(* IEC 61131-3 sources: nautilus/tools/blackbox/projects/2026-10-24-001d/typed, 2 files *)

(* ---- types.st ---- *)
(* library file: types used by the typed project *)
TYPE Mode : (Idle, Run := 10, Fault) := Idle; END_TYPE
TYPE Drive : STRUCT
    Speed : REAL;
    Amps  : REAL;
  END_STRUCT;
END_TYPE
TYPE Motor : STRUCT
    Running : BOOL;
    Fault   : BOOL;
    Starts  : DINT;
    Drive   : Drive;
    State   : Mode;
  END_STRUCT;
END_TYPE
TYPE DoseRecipe : STRUCT
    TargetL    : REAL;
    SettleTime : TIME;
    Steps      : ARRAY[0..2] OF TIME;
  END_STRUCT;
END_TYPE

(* ---- main.st ---- *)
PROGRAM Main
VAR_EXTERNAL
    Counter  : DINT;
    Ramp     : REAL;
    Blink    : BOOL;
    Fixed    : INT;
    P101     : Motor;
    Pumps    : ARRAY[1..2] OF Motor;
    ScanDt   : REAL;
END_VAR
VAR
    t : TON;
END_VAR
Counter := Counter + 1;
Ramp := Ramp + 0.5;
IF Ramp > 100.0 THEN Ramp := 0.0; END_IF;
Fixed := 7;                         (* same value every scan *)
t(IN := NOT t.Q, PT := T#1s);
IF t.Q THEN Blink := NOT Blink; END_IF;
P101.Drive.Speed := Ramp * 10.0;
P101.Starts := Counter;
Pumps[2].Drive.Amps := Ramp;
END_PROGRAM
